(*
SPDX-FileCopyrightText: c 2026 Oleksandr Tiutyk <trofimich@gmail.com>
SPDX-License-Identifier: MIT
License: https://opensource.org/license/mit
*)

(*
Logs the main runner results to ADS and retains a JUnit report.

The owning runner calls the ADS reporter first and the JUnit reporter second at each reporting boundary.
Callback exceptions abort the runner. The JUnit buffer belongs to this instance and its contents are stable
after a successful ReportRunEnd until the next ReportRunStart. Do not copy this instance or reenter its callbacks.
*)

{attribute 'no_assign'}
{attribute 'no_explicit_call' := 'do not call this function block directly'}
FUNCTION_BLOCK MainTestReporter EXTENDS TOF_Testing.AdsLogReporter
VAR_STAT
	// Concrete reporter class name stored separately from the inherited class name.
	{attribute 'hide'}
	_MainReporterClassName : STRING := __POUNAME();
END_VAR
VAR
	// Owns the JUnit buffer for the main runner.
	_JUnitReporter : TOF_Testing.JUnitXmlReporter;
END_VAR

// Provides the concrete report writer class name.
{attribute 'monitoring' := 'call'}
PROPERTY ClassName : REFERENCE TO STRING
GET
ClassName REF= _MainReporterClassName;
END_GET
END_PROPERTY

// Provides the concrete report writer namespace.
{attribute 'monitoring' := 'call'}
PROPERTY NamespaceName : REFERENCE TO STRING
GET
NamespaceName REF= CurrentNamespace.Name;
END_GET
END_PROPERTY

// Reports this instance's storage excluding the dynamic JUnit buffer.
{attribute 'monitoring' := 'call'}
PROPERTY SelfSize : ULINT
GET
SelfSize := XSIZEOF(THIS^);
END_GET
END_PROPERTY

(*
Reports the completed JUnit document's byte count without the terminating zero.

Returns zero until the JUnit reporter has finished writing the document.
*)
{attribute 'monitoring' := 'call'}
PROPERTY JUnitContentLength : UDINT
GET
IF _JUnitReporter.IsReady THEN
	JUnitContentLength := _JUnitReporter.ContentLength;
END_IF
END_GET
END_PROPERTY

(*
Copies up to 1023 ASCII bytes from the completed JUnit document into an IEC string.

Returns an empty string when the report is unavailable or the offset is at or beyond the end.
Also returns an empty string if the byte copy does not complete.
Read in the owning task while callbacks are idle. The returned string is independent of the reporter buffer.

offset — Zero-based byte offset in the document.
*)
METHOD ReadJUnitChunk : STRING(1023)
VAR_INPUT
	offset : UDINT;
END_VAR
VAR
	contentLength : UDINT;
	source : POINTER TO STRING;
	byteCount : UDINT;
	chunkBytes : ARRAY [0..1023] OF BYTE;
	chunkText : POINTER TO STRING(1023);
END_VAR
ReadJUnitChunk := '';
contentLength := JUnitContentLength;

IF offset >= contentLength THEN
	RETURN;
END_IF

source := _JUnitReporter.ContentAddress;

IF source = 0 THEN
	RETURN;
END_IF

// Reserve the last byte for the ASCII string terminator.
byteCount := MIN(contentLength - offset, TO_UDINT(SIZEOF(chunkBytes)) - 1);

IF Tc2_System.MEMCPY(destAddr := ADR(chunkBytes), srcAddr := source + offset, n := byteCount) = byteCount THEN
	chunkBytes[byteCount] := TO_BYTE(TOF_Core.UnsignedInt8.MIN_VALUE);
	chunkText := ADR(chunkBytes);
	ReadJUnitChunk := chunkText^;
END_IF
END_METHOD

(*
Starts ADS logging and opens the new JUnit document.

The JUnit start invalidates the previous document and reuses the allocated buffer.
*)
METHOD ReportRunStart
VAR_INPUT
	testCount : TOF_Core.DINT_LENGTH;
END_VAR
SUPER^.ReportRunStart(testCount := testCount);
_JUnitReporter.ReportRunStart(testCount := testCount);
END_METHOD

(*
Reports a terminal leaf to ADS and adds its testcase to the JUnit document.

Accepts the terminal outcomes defined by ITestReporter. The diagnostic is borrowed for this call.
*)
METHOD ReportTestCaseResult
VAR_INPUT
	groupPath : WSTRING(255);
	testName : WSTRING;
	outcome : TOF_Testing.TEST_OUTCOME;
	duration : TIME;
END_VAR
VAR_IN_OUT CONSTANT
	message : TOF_Core.ERROR_MESSAGE;
END_VAR
SUPER^.ReportTestCaseResult(
	groupPath := groupPath,
	testName := testName,
	outcome := outcome,
	duration := duration,
	message := message
);
_JUnitReporter.ReportTestCaseResult(
	groupPath := groupPath,
	testName := testName,
	outcome := outcome,
	duration := duration,
	message := message
);
END_METHOD

(*
Retains the ADS summary and closes the JUnit document.

After this callback succeeds, both outputs describe the same completed main run.
*)
METHOD ReportRunEnd
VAR_INPUT
	totalTests : TOF_Core.DINT_LENGTH;
	passedTests : TOF_Core.DINT_LENGTH;
	failedTests : TOF_Core.DINT_LENGTH;
	skippedTests : TOF_Core.DINT_LENGTH;
	duration : TIME;
END_VAR
SUPER^.ReportRunEnd(
	totalTests := totalTests,
	passedTests := passedTests,
	failedTests := failedTests,
	skippedTests := skippedTests,
	duration := duration
);
_JUnitReporter.ReportRunEnd(
	totalTests := totalTests,
	passedTests := passedTests,
	failedTests := failedTests,
	skippedTests := skippedTests,
	duration := duration
);
END_METHOD

END_FUNCTION_BLOCK

(* stored: Version 1.1.0.1
   POU MainTestReporter: Id {7eb12daa-2e96-44ac-82a1-0e136171df21}, SpecialFunc None
   Property ClassName: Id {8d7366ea-239d-4c0f-afb1-c02d1f244978}
   Get Get: Id {e3f6574e-9f4b-4980-a8cd-06c64372ab96}
   Property NamespaceName: Id {1ae55fc9-f332-41c1-8c48-6d86650c384f}
   Get Get: Id {a85dbd59-1830-4cda-9643-15a3ab2fafc2}
   Property SelfSize: Id {1c6051a3-88af-4920-9034-dd9f3921eb0e}
   Get Get: Id {971d65b2-9966-4448-9c28-9a2cde9ae5ed}
   Property JUnitContentLength: Id {df140cf5-fd9c-44d1-a577-ae98f247c746}
   Get Get: Id {cf9052f9-5b13-4227-829f-af02bd923279}
   Method ReadJUnitChunk: Id {20ed118a-cd2e-40f3-b3f1-8ccf8a15008d}
   Method ReportRunStart: Id {a35df40e-91a6-42db-9795-e2913ec89978}
   Method ReportTestCaseResult: Id {ef4e5cf7-e97f-49fd-a060-d254781c8a07}
   Method ReportRunEnd: Id {d55cbe5b-1ae1-4ad0-9387-1e57bac6a9c2} *)
